# EPICS autosave request: utcaApp/Db/bpm_pico.req
$(P)$(R)FMCPICORngR0-Sel
$(P)$(R)FMCPICORngR1-Sel
$(P)$(R)FMCPICORngR2-Sel
$(P)$(R)FMCPICORngR3-Sel
